Yaskawa INFORM job: 4043MMR1.JBI

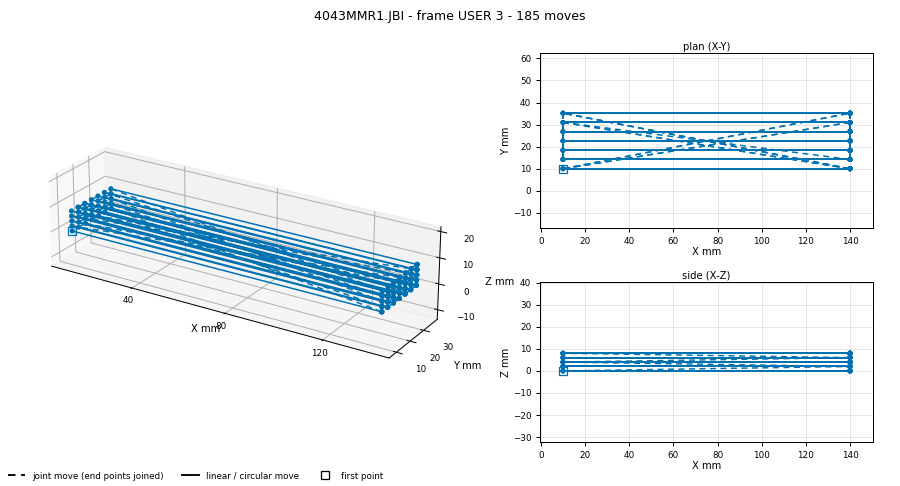
[picture p0: tool path of 4043MMR1.JBI in frame USER 3, 185 of 185 moves have a stored position in this frame; points joined in program order, loops and branches not executed]
/JOB
//NAME 4043MMR1
//POS
///NPOS 185,0,0,0,0,0
///USER 3
///TOOL 1
///POSTYPE USER
///RECTAN
///RCONF 1,0,0,0,0,0,0,0,0,0,0,0,0,0,0,0,0,0,0,0,0,0,0,0
C00000=10.000,10.000,0.000,0.0000,0.0000,-110.0000
C00001=140.000,10.000,0.000,0.0000,0.0000,-110.0000
C00002=140.000,10.000,0.000,0.0000,0.0000,-110.0000
C00003=140.000,10.000,0.000,0.0000,0.0000,-110.0000
C00004=140.000,10.000,0.000,0.0000,0.0000,-110.0000
C00005=10.000,35.200,0.000,0.0000,0.0000,-110.0000
C00006=140.000,35.200,0.000,0.0000,0.0000,-110.0000
C00007=140.000,35.200,0.000,0.0000,0.0000,-110.0000
C00008=140.000,35.200,0.000,0.0000,0.0000,-110.0000
C00009=140.000,35.200,0.000,0.0000,0.0000,-110.0000
C00010=140.000,14.200,0.000,0.0000,0.0000,-110.0000
C00011=140.000,14.200,0.000,0.0000,0.0000,-110.0000
C00012=140.000,14.200,0.000,0.0000,0.0000,-110.0000
C00013=140.000,14.200,0.000,0.0000,0.0000,-110.0000
C00014=10.000,14.200,0.000,0.0000,0.0000,-110.0000
C00015=10.000,18.400,0.000,0.0000,0.0000,-110.0000
C00016=140.000,18.400,0.000,0.0000,0.0000,-110.0000
C00017=140.000,18.400,0.000,0.0000,0.0000,-110.0000
C00018=140.000,18.400,0.000,0.0000,0.0000,-110.0000
C00019=140.000,18.400,0.000,0.0000,0.0000,-110.0000
C00020=140.000,22.600,0.000,0.0000,0.0000,-110.0000
C00021=140.000,22.600,0.000,0.0000,0.0000,-110.0000
C00022=140.000,22.600,0.000,0.0000,0.0000,-110.0000
C00023=140.000,22.600,0.000,0.0000,0.0000,-110.0000
C00024=10.000,22.600,0.000,0.0000,0.0000,-110.0000
C00025=10.000,26.800,0.000,0.0000,0.0000,-110.0000
C00026=140.000,26.800,0.000,0.0000,0.0000,-110.0000
C00027=140.000,26.800,0.000,0.0000,0.0000,-110.0000
C00028=140.000,26.800,0.000,0.0000,0.0000,-110.0000
C00029=140.000,26.800,0.000,0.0000,0.0000,-110.0000
C00030=140.000,31.000,0.000,0.0000,0.0000,-110.0000
C00031=140.000,31.000,0.000,0.0000,0.0000,-110.0000
C00032=140.000,31.000,0.000,0.0000,0.0000,-110.0000
C00033=140.000,31.000,0.000,0.0000,0.0000,-110.0000
C00034=10.000,31.000,0.000,0.0000,0.0000,-110.0000
C00035=140.000,10.000,2.000,0.0000,0.0000,-110.0000
C00036=140.000,10.000,2.000,0.0000,0.0000,-110.0000
C00037=140.000,10.000,2.000,0.0000,0.0000,-110.0000
C00038=140.000,10.000,2.000,0.0000,0.0000,-110.0000
C00039=10.000,10.000,2.000,0.0000,0.0000,-110.0000
C00040=140.000,35.200,2.000,0.0000,0.0000,-110.0000
C00041=140.000,35.200,2.000,0.0000,0.0000,-110.0000
C00042=140.000,35.200,2.000,0.0000,0.0000,-110.0000
C00043=140.000,35.200,2.000,0.0000,0.0000,-110.0000
C00044=10.000,35.200,2.000,0.0000,0.0000,-110.0000
C00045=10.000,14.200,2.000,0.0000,0.0000,-110.0000
C00046=140.000,14.200,2.000,0.0000,0.0000,-110.0000
C00047=140.000,14.200,2.000,0.0000,0.0000,-110.0000
C00048=140.000,14.200,2.000,0.0000,0.0000,-110.0000
C00049=140.000,14.200,2.000,0.0000,0.0000,-110.0000
C00050=140.000,18.400,2.000,0.0000,0.0000,-110.0000
C00051=140.000,18.400,2.000,0.0000,0.0000,-110.0000
C00052=140.000,18.400,2.000,0.0000,0.0000,-110.0000
C00053=140.000,18.400,2.000,0.0000,0.0000,-110.0000
C00054=10.000,18.400,2.000,0.0000,0.0000,-110.0000
C00055=10.000,22.600,2.000,0.0000,0.0000,-110.0000
C00056=140.000,22.600,2.000,0.0000,0.0000,-110.0000
C00057=140.000,22.600,2.000,0.0000,0.0000,-110.0000
C00058=140.000,22.600,2.000,0.0000,0.0000,-110.0000
C00059=140.000,22.600,2.000,0.0000,0.0000,-110.0000
C00060=140.000,26.800,2.000,0.0000,0.0000,-110.0000
C00061=140.000,26.800,2.000,0.0000,0.0000,-110.0000
C00062=140.000,26.800,2.000,0.0000,0.0000,-110.0000
C00063=140.000,26.800,2.000,0.0000,0.0000,-110.0000
C00064=10.000,26.800,2.000,0.0000,0.0000,-110.0000
C00065=10.000,31.000,2.000,0.0000,0.0000,-110.0000
C00066=140.000,31.000,2.000,0.0000,0.0000,-110.0000
C00067=140.000,31.000,2.000,0.0000,0.0000,-110.0000
C00068=140.000,31.000,2.000,0.0000,0.0000,-110.0000
C00069=140.000,31.000,2.000,0.0000,0.0000,-110.0000
C00070=10.000,10.000,4.000,0.0000,0.0000,-110.0000
C00071=140.000,10.000,4.000,0.0000,0.0000,-110.0000
C00072=140.000,10.000,4.000,0.0000,0.0000,-110.0000
C00073=140.000,10.000,4.000,0.0000,0.0000,-110.0000
C00074=140.000,10.000,4.000,0.0000,0.0000,-110.0000
C00075=10.000,35.200,4.000,0.0000,0.0000,-110.0000
C00076=140.000,35.200,4.000,0.0000,0.0000,-110.0000
C00077=140.000,35.200,4.000,0.0000,0.0000,-110.0000
C00078=140.000,35.200,4.000,0.0000,0.0000,-110.0000
C00079=140.000,35.200,4.000,0.0000,0.0000,-110.0000
C00080=140.000,14.200,4.000,0.0000,0.0000,-110.0000
C00081=140.000,14.200,4.000,0.0000,0.0000,-110.0000
C00082=140.000,14.200,4.000,0.0000,0.0000,-110.0000
C00083=140.000,14.200,4.000,0.0000,0.0000,-110.0000
C00084=10.000,14.200,4.000,0.0000,0.0000,-110.0000
C00085=10.000,18.400,4.000,0.0000,0.0000,-110.0000
C00086=140.000,18.400,4.000,0.0000,0.0000,-110.0000
C00087=140.000,18.400,4.000,0.0000,0.0000,-110.0000
C00088=140.000,18.400,4.000,0.0000,0.0000,-110.0000
C00089=140.000,18.400,4.000,0.0000,0.0000,-110.0000
C00090=140.000,22.600,4.000,0.0000,0.0000,-110.0000
C00091=140.000,22.600,4.000,0.0000,0.0000,-110.0000
C00092=140.000,22.600,4.000,0.0000,0.0000,-110.0000
C00093=140.000,22.600,4.000,0.0000,0.0000,-110.0000
C00094=10.000,22.600,4.000,0.0000,0.0000,-110.0000
C00095=10.000,26.800,4.000,0.0000,0.0000,-110.0000
C00096=140.000,26.800,4.000,0.0000,0.0000,-110.0000
C00097=140.000,26.800,4.000,0.0000,0.0000,-110.0000
C00098=140.000,26.800,4.000,0.0000,0.0000,-110.0000
C00099=140.000,26.800,4.000,0.0000,0.0000,-110.0000
C00100=140.000,31.000,4.000,0.0000,0.0000,-110.0000
C00101=140.000,31.000,4.000,0.0000,0.0000,-110.0000
C00102=140.000,31.000,4.000,0.0000,0.0000,-110.0000
C00103=140.000,31.000,4.000,0.0000,0.0000,-110.0000
C00104=10.000,31.000,4.000,0.0000,0.0000,-110.0000
C00105=140.000,10.000,6.000,0.0000,0.0000,-110.0000
C00106=140.000,10.000,6.000,0.0000,0.0000,-110.0000
C00107=140.000,10.000,6.000,0.0000,0.0000,-110.0000
C00108=140.000,10.000,6.000,0.0000,0.0000,-110.0000
C00109=10.000,10.000,6.000,0.0000,0.0000,-110.0000
C00110=140.000,35.200,6.000,0.0000,0.0000,-110.0000
C00111=140.000,35.200,6.000,0.0000,0.0000,-110.0000
C00112=140.000,35.200,6.000,0.0000,0.0000,-110.0000
C00113=140.000,35.200,6.000,0.0000,0.0000,-110.0000
C00114=10.000,35.200,6.000,0.0000,0.0000,-110.0000
C00115=10.000,14.200,6.000,0.0000,0.0000,-110.0000
C00116=140.000,14.200,6.000,0.0000,0.0000,-110.0000
C00117=140.000,14.200,6.000,0.0000,0.0000,-110.0000
C00118=140.000,14.200,6.000,0.0000,0.0000,-110.0000
C00119=140.000,14.200,6.000,0.0000,0.0000,-110.0000
C00120=140.000,18.400,6.000,0.0000,0.0000,-110.0000
C00121=140.000,18.400,6.000,0.0000,0.0000,-110.0000
C00122=140.000,18.400,6.000,0.0000,0.0000,-110.0000
C00123=140.000,18.400,6.000,0.0000,0.0000,-110.0000
C00124=10.000,18.400,6.000,0.0000,0.0000,-110.0000
C00125=10.000,22.600,6.000,0.0000,0.0000,-110.0000
C00126=140.000,22.600,6.000,0.0000,0.0000,-110.0000
C00127=140.000,22.600,6.000,0.0000,0.0000,-110.0000
C00128=140.000,22.600,6.000,0.0000,0.0000,-110.0000
C00129=140.000,22.600,6.000,0.0000,0.0000,-110.0000
C00130=140.000,26.800,6.000,0.0000,0.0000,-110.0000
C00131=140.000,26.800,6.000,0.0000,0.0000,-110.0000
C00132=140.000,26.800,6.000,0.0000,0.0000,-110.0000
C00133=140.000,26.800,6.000,0.0000,0.0000,-110.0000
C00134=10.000,26.800,6.000,0.0000,0.0000,-110.0000
C00135=10.000,31.000,6.000,0.0000,0.0000,-110.0000
C00136=140.000,31.000,6.000,0.0000,0.0000,-110.0000
C00137=140.000,31.000,6.000,0.0000,0.0000,-110.0000
C00138=140.000,31.000,6.000,0.0000,0.0000,-110.0000
C00139=140.000,31.000,6.000,0.0000,0.0000,-110.0000
C00140=10.000,10.000,8.000,0.0000,0.0000,-110.0000
C00141=140.000,10.000,8.000,0.0000,0.0000,-110.0000
C00142=140.000,10.000,8.000,0.0000,0.0000,-110.0000
C00143=140.000,10.000,8.000,0.0000,0.0000,-110.0000
C00144=140.000,10.000,8.000,0.0000,0.0000,-110.0000
C00145=10.000,35.200,8.000,0.0000,0.0000,-110.0000
C00146=140.000,35.200,8.000,0.0000,0.0000,-110.0000
C00147=140.000,35.200,8.000,0.0000,0.0000,-110.0000
C00148=140.000,35.200,8.000,0.0000,0.0000,-110.0000
C00149=140.000,35.200,8.000,0.0000,0.0000,-110.0000
C00150=140.000,14.200,8.000,0.0000,0.0000,-110.0000
C00151=140.000,14.200,8.000,0.0000,0.0000,-110.0000
C00152=140.000,14.200,8.000,0.0000,0.0000,-110.0000
C00153=140.000,14.200,8.000,0.0000,0.0000,-110.0000
C00154=10.000,14.200,8.000,0.0000,0.0000,-110.0000
C00155=10.000,18.400,8.000,0.0000,0.0000,-110.0000
C00156=140.000,18.400,8.000,0.0000,0.0000,-110.0000
C00157=140.000,18.400,8.000,0.0000,0.0000,-110.0000
C00158=140.000,18.400,8.000,0.0000,0.0000,-110.0000
C00159=140.000,18.400,8.000,0.0000,0.0000,-110.0000
C00160=140.000,22.600,8.000,0.0000,0.0000,-110.0000
C00161=140.000,22.600,8.000,0.0000,0.0000,-110.0000
C00162=140.000,22.600,8.000,0.0000,0.0000,-110.0000
C00163=140.000,22.600,8.000,0.0000,0.0000,-110.0000
C00164=10.000,22.600,8.000,0.0000,0.0000,-110.0000
C00165=10.000,26.800,8.000,0.0000,0.0000,-110.0000
C00166=140.000,26.800,8.000,0.0000,0.0000,-110.0000
C00167=140.000,26.800,8.000,0.0000,0.0000,-110.0000
C00168=140.000,26.800,8.000,0.0000,0.0000,-110.0000
C00169=140.000,26.800,8.000,0.0000,0.0000,-110.0000
C00170=140.000,31.000,8.000,0.0000,0.0000,-110.0000
C00171=140.000,31.000,8.000,0.0000,0.0000,-110.0000
C00172=140.000,31.000,8.000,0.0000,0.0000,-110.0000
C00173=140.000,31.000,8.000,0.0000,0.0000,-110.0000
C00174=10.000,31.000,8.000,0.0000,0.0000,-110.0000
C00175=140.000,14.200,8.000,0.0000,0.0000,-110.0000
C00176=140.000,14.200,8.000,0.0000,0.0000,-110.0000
C00177=140.000,14.200,8.000,0.0000,0.0000,-110.0000
C00178=140.000,14.200,8.000,0.0000,0.0000,-110.0000
C00179=10.000,14.200,8.000,0.0000,0.0000,-110.0000
C00180=10.000,18.400,8.000,0.0000,0.0000,-110.0000
C00181=140.000,18.400,8.000,0.0000,0.0000,-110.0000
C00182=140.000,18.400,8.000,0.0000,0.0000,-110.0000
C00183=140.000,18.400,8.000,0.0000,0.0000,-110.0000
C00184=140.000,18.400,8.000,0.0000,0.0000,-110.0000
//INST
///DATE 2025/03/17 13:38
///COMM Grasshopper
///ATTR SC,RW,RJ
////FRAME USER 3
///GROUP1 RB1
NOP
DOUT OT#(9) OFF
TIMER T=5.00
*LABEL0
MOVJ C00000 VJ=10.00 ACC=20
MACRO1 MJ#(0) ARGF200
ARCON
MOVL C00001 V=12.0 ACC=20
MOVL C00002 V=12.0 ACC=20
MOVL C00003 V=12.0 ACC=20
MOVL C00004 V=12.0 ACC=20
ARCOF
TIMER T=7.00
*LABEL1
MOVJ C00005 VJ=10.00 ACC=20
MACRO1 MJ#(0) ARGF200
ARCON
MOVL C00006 V=12.0 ACC=20
MOVL C00007 V=12.0 ACC=20
MOVL C00008 V=12.0 ACC=20
MOVL C00009 V=12.0 ACC=20
ARCOF
DOUT OT#(9) ON
TIMER T=50.00
DOUT OT#(9) OFF
TIMER T=13.00
*LABEL2
MOVJ C00010 VJ=10.00 ACC=20
MACRO1 MJ#(0) ARGF200
ARCON
MOVL C00011 V=12.0 ACC=20
MOVL C00012 V=12.0 ACC=20
MOVL C00013 V=12.0 ACC=20
MOVL C00014 V=12.0 ACC=20
ARCOF
TIMER T=7.00
*LABEL3
MOVJ C00015 VJ=10.00 ACC=20
MACRO1 MJ#(0) ARGF200
ARCON
MOVL C00016 V=12.0 ACC=20
MOVL C00017 V=12.0 ACC=20
MOVL C00018 V=12.0 ACC=20
MOVL C00019 V=12.0 ACC=20
ARCOF
TIMER T=7.00
*LABEL4
MOVJ C00020 VJ=10.00 ACC=20
MACRO1 MJ#(0) ARGF200
ARCON
MOVL C00021 V=12.0 ACC=20
MOVL C00022 V=12.0 ACC=20
MOVL C00023 V=12.0 ACC=20
MOVL C00024 V=12.0 ACC=20
ARCOF
TIMER T=7.00
*LABEL5
MOVJ C00025 VJ=10.00 ACC=20
MACRO1 MJ#(0) ARGF200
ARCON
MOVL C00026 V=12.0 ACC=20
MOVL C00027 V=12.0 ACC=20
MOVL C00028 V=12.0 ACC=20
MOVL C00029 V=12.0 ACC=20
ARCOF
TIMER T=7.00
*LABEL6
MOVJ C00030 VJ=10.00 ACC=20
MACRO1 MJ#(0) ARGF200
ARCON
MOVL C00031 V=12.0 ACC=20
MOVL C00032 V=12.0 ACC=20
MOVL C00033 V=12.0 ACC=20
MOVL C00034 V=12.0 ACC=20
ARCOF
DOUT OT#(9) ON
TIMER T=50.00
DOUT OT#(9) OFF
TIMER T=13.00
*LABEL7
MOVJ C00035 VJ=10.00 ACC=20
MACRO1 MJ#(0) ARGF200
ARCON
MOVL C00036 V=12.0 ACC=20
MOVL C00037 V=12.0 ACC=20
MOVL C00038 V=12.0 ACC=20
MOVL C00039 V=12.0 ACC=20
ARCOF
TIMER T=7.00
*LABEL8
MOVJ C00040 VJ=10.00 ACC=20
MACRO1 MJ#(0) ARGF200
ARCON
MOVL C00041 V=12.0 ACC=20
MOVL C00042 V=12.0 ACC=20
MOVL C00043 V=12.0 ACC=20
MOVL C00044 V=12.0 ACC=20
ARCOF
DOUT OT#(9) ON
TIMER T=50.00
DOUT OT#(9) OFF
TIMER T=13.00
*LABEL9
MOVJ C00045 VJ=10.00 ACC=20
MACRO1 MJ#(0) ARGF200
ARCON
MOVL C00046 V=12.0 ACC=20
MOVL C00047 V=12.0 ACC=20
MOVL C00048 V=12.0 ACC=20
MOVL C00049 V=12.0 ACC=20
ARCOF
TIMER T=7.00
*LABEL10
MOVJ C00050 VJ=10.00 ACC=20
MACRO1 MJ#(0) ARGF200
ARCON
MOVL C00051 V=12.0 ACC=20
MOVL C00052 V=12.0 ACC=20
MOVL C00053 V=12.0 ACC=20
MOVL C00054 V=12.0 ACC=20
ARCOF
TIMER T=7.00
*LABEL11
MOVJ C00055 VJ=10.00 ACC=20
MACRO1 MJ#(0) ARGF200
ARCON
MOVL C00056 V=12.0 ACC=20
MOVL C00057 V=12.0 ACC=20
MOVL C00058 V=12.0 ACC=20
MOVL C00059 V=12.0 ACC=20
ARCOF
TIMER T=7.00
*LABEL12
MOVJ C00060 VJ=10.00 ACC=20
MACRO1 MJ#(0) ARGF200
ARCON
MOVL C00061 V=12.0 ACC=20
MOVL C00062 V=12.0 ACC=20
MOVL C00063 V=12.0 ACC=20
MOVL C00064 V=12.0 ACC=20
ARCOF
TIMER T=7.00
*LABEL13
MOVJ C00065 VJ=10.00 ACC=20
MACRO1 MJ#(0) ARGF200
ARCON
MOVL C00066 V=12.0 ACC=20
MOVL C00067 V=12.0 ACC=20
MOVL C00068 V=12.0 ACC=20
MOVL C00069 V=12.0 ACC=20
ARCOF
DOUT OT#(9) ON
TIMER T=50.00
DOUT OT#(9) OFF
TIMER T=13.00
*LABEL14
MOVJ C00070 VJ=10.00 ACC=20
MACRO1 MJ#(0) ARGF200
ARCON
MOVL C00071 V=12.0 ACC=20
MOVL C00072 V=12.0 ACC=20
MOVL C00073 V=12.0 ACC=20
MOVL C00074 V=12.0 ACC=20
ARCOF
TIMER T=7.00
*LABEL15
MOVJ C00075 VJ=10.00 ACC=20
MACRO1 MJ#(0) ARGF200
ARCON
MOVL C00076 V=12.0 ACC=20
MOVL C00077 V=12.0 ACC=20
MOVL C00078 V=12.0 ACC=20
MOVL C00079 V=12.0 ACC=20
ARCOF
DOUT OT#(9) ON
TIMER T=50.00
DOUT OT#(9) OFF
TIMER T=13.00
*LABEL16
MOVJ C00080 VJ=10.00 ACC=20
MACRO1 MJ#(0) ARGF200
ARCON
MOVL C00081 V=12.0 ACC=20
MOVL C00082 V=12.0 ACC=20
MOVL C00083 V=12.0 ACC=20
MOVL C00084 V=12.0 ACC=20
ARCOF
TIMER T=7.00
*LABEL17
MOVJ C00085 VJ=10.00 ACC=20
MACRO1 MJ#(0) ARGF200
ARCON
MOVL C00086 V=12.0 ACC=20
MOVL C00087 V=12.0 ACC=20
MOVL C00088 V=12.0 ACC=20
MOVL C00089 V=12.0 ACC=20
ARCOF
TIMER T=7.00
*LABEL18
MOVJ C00090 VJ=10.00 ACC=20
MACRO1 MJ#(0) ARGF200
ARCON
MOVL C00091 V=12.0 ACC=20
MOVL C00092 V=12.0 ACC=20
MOVL C00093 V=12.0 ACC=20
MOVL C00094 V=12.0 ACC=20
ARCOF
TIMER T=7.00
*LABEL19
MOVJ C00095 VJ=10.00 ACC=20
MACRO1 MJ#(0) ARGF200
ARCON
MOVL C00096 V=12.0 ACC=20
MOVL C00097 V=12.0 ACC=20
MOVL C00098 V=12.0 ACC=20
MOVL C00099 V=12.0 ACC=20
ARCOF
TIMER T=7.00
*LABEL20
MOVJ C00100 VJ=10.00 ACC=20
MACRO1 MJ#(0) ARGF200
ARCON
MOVL C00101 V=12.0 ACC=20
MOVL C00102 V=12.0 ACC=20
MOVL C00103 V=12.0 ACC=20
MOVL C00104 V=12.0 ACC=20
ARCOF
DOUT OT#(9) ON
TIMER T=50.00
DOUT OT#(9) OFF
TIMER T=13.00
*LABEL21
MOVJ C00105 VJ=10.00 ACC=20
MACRO1 MJ#(0) ARGF200
ARCON
MOVL C00106 V=12.0 ACC=20
MOVL C00107 V=12.0 ACC=20
MOVL C00108 V=12.0 ACC=20
MOVL C00109 V=12.0 ACC=20
ARCOF
TIMER T=7.00
*LABEL22
MOVJ C00110 VJ=10.00 ACC=20
MACRO1 MJ#(0) ARGF200
ARCON
MOVL C00111 V=12.0 ACC=20
MOVL C00112 V=12.0 ACC=20
MOVL C00113 V=12.0 ACC=20
MOVL C00114 V=12.0 ACC=20
ARCOF
DOUT OT#(9) ON
TIMER T=50.00
DOUT OT#(9) OFF
TIMER T=13.00
*LABEL23
MOVJ C00115 VJ=10.00 ACC=20
MACRO1 MJ#(0) ARGF200
ARCON
MOVL C00116 V=12.0 ACC=20
MOVL C00117 V=12.0 ACC=20
MOVL C00118 V=12.0 ACC=20
MOVL C00119 V=12.0 ACC=20
ARCOF
TIMER T=7.00
*LABEL24
MOVJ C00120 VJ=10.00 ACC=20
MACRO1 MJ#(0) ARGF200
ARCON
MOVL C00121 V=12.0 ACC=20
MOVL C00122 V=12.0 ACC=20
MOVL C00123 V=12.0 ACC=20
MOVL C00124 V=12.0 ACC=20
ARCOF
TIMER T=7.00
*LABEL25
MOVJ C00125 VJ=10.00 ACC=20
MACRO1 MJ#(0) ARGF200
ARCON
MOVL C00126 V=12.0 ACC=20
MOVL C00127 V=12.0 ACC=20
MOVL C00128 V=12.0 ACC=20
MOVL C00129 V=12.0 ACC=20
ARCOF
TIMER T=7.00
*LABEL26
MOVJ C00130 VJ=10.00 ACC=20
MACRO1 MJ#(0) ARGF200
ARCON
MOVL C00131 V=12.0 ACC=20
MOVL C00132 V=12.0 ACC=20
MOVL C00133 V=12.0 ACC=20
MOVL C00134 V=12.0 ACC=20
ARCOF
TIMER T=7.00
*LABEL27
MOVJ C00135 VJ=10.00 ACC=20
MACRO1 MJ#(0) ARGF200
ARCON
MOVL C00136 V=12.0 ACC=20
MOVL C00137 V=12.0 ACC=20
MOVL C00138 V=12.0 ACC=20
MOVL C00139 V=12.0 ACC=20
ARCOF
DOUT OT#(9) ON
TIMER T=50.00
DOUT OT#(9) OFF
TIMER T=13.00
*LABEL28
MOVJ C00140 VJ=10.00 ACC=20
MACRO1 MJ#(0) ARGF200
ARCON
MOVL C00141 V=12.0 ACC=20
MOVL C00142 V=12.0 ACC=20
MOVL C00143 V=12.0 ACC=20
MOVL C00144 V=12.0 ACC=20
ARCOF
TIMER T=7.00
*LABEL29
MOVJ C00145 VJ=10.00 ACC=20
MACRO1 MJ#(0) ARGF200
ARCON
MOVL C00146 V=12.0 ACC=20
MOVL C00147 V=12.0 ACC=20
MOVL C00148 V=12.0 ACC=20
MOVL C00149 V=12.0 ACC=20
ARCOF
DOUT OT#(9) ON
TIMER T=50.00
DOUT OT#(9) OFF
TIMER T=13.00
*LABEL30
MOVJ C00150 VJ=10.00 ACC=20
MACRO1 MJ#(0) ARGF200
ARCON
MOVL C00151 V=12.0 ACC=20
MOVL C00152 V=12.0 ACC=20
MOVL C00153 V=12.0 ACC=20
MOVL C00154 V=12.0 ACC=20
ARCOF
TIMER T=7.00
*LABEL31
MOVJ C00155 VJ=10.00 ACC=20
MACRO1 MJ#(0) ARGF200
ARCON
MOVL C00156 V=12.0 ACC=20
MOVL C00157 V=12.0 ACC=20
MOVL C00158 V=12.0 ACC=20
MOVL C00159 V=12.0 ACC=20
ARCOF
TIMER T=7.00
*LABEL32
MOVJ C00160 VJ=10.00 ACC=20
MACRO1 MJ#(0) ARGF200
ARCON
MOVL C00161 V=12.0 ACC=20
MOVL C00162 V=12.0 ACC=20
MOVL C00163 V=12.0 ACC=20
MOVL C00164 V=12.0 ACC=20
ARCOF
TIMER T=7.00
*LABEL33
MOVJ C00165 VJ=10.00 ACC=20
MACRO1 MJ#(0) ARGF200
ARCON
MOVL C00166 V=12.0 ACC=20
MOVL C00167 V=12.0 ACC=20
MOVL C00168 V=12.0 ACC=20
MOVL C00169 V=12.0 ACC=20
ARCOF
TIMER T=7.00
*LABEL34
MOVJ C00170 VJ=10.00 ACC=20
MACRO1 MJ#(0) ARGF200
ARCON
MOVL C00171 V=12.0 ACC=20
MOVL C00172 V=12.0 ACC=20
MOVL C00173 V=12.0 ACC=20
MOVL C00174 V=12.0 ACC=20
ARCOF
DOUT OT#(9) ON
TIMER T=50.00
DOUT OT#(9) OFF
TIMER T=13.00
JUMP *LABEL34E
JUMP *LABEL999
*LABEL34E
MOVJ C00175 VJ=10.00 ACC=20
MACRO1 MJ#(0) ARGF103
ARCON
MOVL C00176 V=12.0 ACC=20
MOVL C00177 V=12.0 ACC=20
MOVL C00178 V=12.0 ACC=20
MOVL C00179 V=12.0 ACC=20
ARCOF
TIMER T=7.00
MOVJ C00180 VJ=10.00 ACC=20
MACRO1 MJ#(0) ARGF103
ARCON
MOVL C00181 V=12.0 ACC=20
MOVL C00182 V=12.0 ACC=20
MOVL C00183 V=12.0 ACC=20
MOVL C00184 V=12.0 ACC=20
ARCOF
DOUT OT#(9) ON
TIMER T=50.00
DOUT OT#(9) OFF
TIMER T=13.00
*LABEL999
END
